VAR_GLOBAL
	(* values of the pointing model
	Hour Angle	: tau
	Declination	: dec
	*)

	(*
	 pointing from: 21.01.2026 136 points (from Lukas Melzig)
	RMS Ha:  17.69244750276253
	RMS Dec:  13.468555776826959
	*)
	C_mAl_tau	: LREAL := 0.01687078;
	C_mEl_tau	: LREAL := -0.02608578;
	C_Coll_tau	: LREAL := 0.29826615;
	C_Refr_tau	: LREAL := -0.00759962;
	C_Enc_tau	: LREAL := 0.00108764;
	C_Flex_tau	: LREAL := -0.02462705;
	C_NP_tau	: LREAL := 0.02128217;
	
	C_mAl_dec	: LREAL := 0.01606325;
	C_mEl_dec	: LREAL := -0.05749048;
	C_Coll_dec	: LREAL := -0.17376101;
	C_Refr_dec	: LREAL := 0.01678090;
	C_Flex_dec	: LREAL := -0.01915146;
END_VAR

(* stored: Version 1.1.0.1, ProductVersion 3.1.4024.15
   GVL GVL_Pointing: Id {8e9e0956-bbc2-49ba-acc4-8eac020b70e3} *)
